(* IEC 61131-3 sources: TetherPLC/tests/ops/cases, 40 files *)

(* ---- o01_debounce.st ---- *)
// o01_debounce.st — FB_AtcDebounce: OnTime=0.3 s sets Q, OffTime=0.2 s
// resets it, ct=0.1 s/scan. D high at n=1 -> Q at n=3 (0.3 s).
// D low at n=6 -> Q clears at n=7 (0.2 s). ET counts since change.
// Sticky bits -> flags %QB0: b0 Q set, b1 Q cleared, b2 ET sane.
PROGRAM O01
VAR
    flags AT %QB0 : BYTE;
    ok0, ok1, ok2 : BOOL;
    deb : FB_AtcDebounce;
    d : BOOL;
    n : DINT;
END_VAR
    n := n + 1;
    IF n = 1 THEN d := TRUE; END_IF;
    IF n = 6 THEN d := FALSE; END_IF;
    deb(D := d, OnTime := 0.3, OffTime := 0.2, CycleTime := 0.1);
    IF n >= 3 AND n < 6 AND deb.Q THEN ok0 := TRUE; END_IF;
    IF n >= 7 AND NOT deb.Q AND n < 30 THEN ok1 := TRUE; END_IF;
    IF n >= 10 AND n < 30 AND deb.ET > 0.05 THEN ok2 := TRUE; END_IF;
    flags := 0;
    IF ok0 THEN flags := flags + 1; END_IF;
    IF ok1 THEN flags := flags + 2; END_IF;
    IF ok2 THEN flags := flags + 4; END_IF;
END_PROGRAM

(* ---- o02_alarm.st ---- *)
// o02_alarm.st — FB_AtcAlarm: Cond edge latches Unacked (survives
// Cond clear), Ack clears it, Shelve suppresses Active for
// ShelveTime s, FirstOut respects HigherPriActive.
//   n=1 Cond up   -> Active+Unacked, FirstOut (no higher pri)
//   n=2 Cond down -> Unacked stays, Active off
//   n=3 Ack       -> Unacked off
//   n=4 Cond up   -> edge again (ack still held -> net unacked off)
//   n=5 Shelve 1s -> Active off, Shelved on
//   n=6..13 shelf window: alm2 (same cond, no shelve, higher-pri =
//        alm.Active=FALSE) -> FirstOut TRUE while alm suppressed
//   n=15+ shelf expires -> alm Active back -> alm2 FirstOut off
// Sticky: b0 unacked latch, b1 ack clears, b2 shelve works,
// b3 shelf expiry restores, b4 firstout suppression.
PROGRAM O02
VAR
    flags AT %QB0 : BYTE;
    ok0, ok1, ok2, ok3, ok4 : BOOL;
    alm : FB_AtcAlarm;
    alm2 : FB_AtcAlarm;
    cond, ack, shelve : BOOL;
    n : DINT;
END_VAR
    n := n + 1;
    IF n = 1 THEN cond := TRUE; END_IF;
    IF n = 2 THEN cond := FALSE; END_IF;
    IF n = 3 THEN ack := TRUE; END_IF;
    IF n = 4 THEN cond := TRUE; END_IF;
    IF n = 5 THEN shelve := TRUE; ack := FALSE; END_IF;
    IF n = 6 THEN shelve := FALSE; END_IF;
    alm(Cond := cond, Ack := ack, Shelve := shelve,
        ShelveTime := 1.0, HigherPriActive := FALSE,
        CycleTime := 0.1);
    alm2(Cond := cond, Ack := FALSE, Shelve := FALSE,
         ShelveTime := 1.0, HigherPriActive := alm.Active,
         CycleTime := 0.1);
    // b0: unacked latched at n=2 even though cond cleared
    IF n = 2 AND alm.Unacked AND NOT alm.Active THEN ok0 := TRUE; END_IF;
    // b1: ack at n=3 cleared unacked
    IF n = 3 AND NOT alm.Unacked THEN ok1 := TRUE; END_IF;
    // b2: shelved at n=6 — cond up but Active suppressed
    IF n = 6 AND alm.Shelved AND NOT alm.Active AND alm.ShelfET > 0.5
       THEN ok2 := TRUE; END_IF;
    // b3: shelf expired -> Active again while cond still up
    IF n >= 15 AND alm.Active AND NOT alm.Shelved THEN ok3 := TRUE; END_IF;
    // b4: during shelf window alm2 is the first-out (alm suppressed)
    IF n = 8 AND alm2.FirstOut AND NOT alm.Active THEN ok4 := TRUE; END_IF;
    flags := 0;
    IF ok0 THEN flags := flags + 1; END_IF;
    IF ok1 THEN flags := flags + 2; END_IF;
    IF ok2 THEN flags := flags + 4; END_IF;
    IF ok3 THEN flags := flags + 8; END_IF;
    IF ok4 THEN flags := flags + 16; END_IF;
END_PROGRAM

(* ---- o03_hourmeter.st ---- *)
// o03_hourmeter.st — FB_AtcHourMeter: ct=3600 s/scan so each scan is
// one hour. Run scans 1-3 -> Hours=3.0, Preset=2.5 -> Alarm + Pct=120.
// Run off at n=4 (hours hold), Reset at n=6 -> zeroed.
// Sticky: b0 hours accumulate, b1 alarm+pct, b2 reset clears.
PROGRAM O03
VAR
    flags AT %QB0 : BYTE;
    ok0, ok1, ok2 : BOOL;
    hm : FB_AtcHourMeter;
    run, rst : BOOL;
    n : DINT;
END_VAR
    n := n + 1;
    run := n <= 3;
    IF n = 6 THEN rst := TRUE; END_IF;
    hm(Run := run, CycleTime := 3600.0, Preset := 2.5, Reset := rst);
    IF n = 3 AND hm.Hours > 2.9 AND hm.Hours < 3.1 THEN ok0 := TRUE; END_IF;
    IF n = 4 AND hm.Alarm AND hm.Pct > 110.0 THEN ok1 := TRUE; END_IF;
    IF n = 7 AND hm.Hours = 0.0 AND NOT hm.Alarm THEN ok2 := TRUE; END_IF;
    flags := 0;
    IF ok0 THEN flags := flags + 1; END_IF;
    IF ok1 THEN flags := flags + 2; END_IF;
    IF ok2 THEN flags := flags + 4; END_IF;
END_PROGRAM

(* ---- o04_oee.st ---- *)
// o04_oee.st — FB_AtcOee: ct=3600 -> 1 h/scan. Planned+Running all
// scans; IdealCycle=10 s. GoodPart pulse n=1, TotalPart pulses n=1,2.
// After n=2: A=100, P=10/(2*3600)*100=0.139, Q=50, OEE~0.069.
// n=8 Reset -> all counters zero, A back to 0 (no plan time).
// Sticky: b0 availability 100, b1 quality 50, b2 perf in band,
// b3 oee in band, b4 reset.
PROGRAM O04
VAR
    flags AT %QB0 : BYTE;
    ok0, ok1, ok2, ok3, ok4 : BOOL;
    oee : FB_AtcOee;
    good, tot, rst : BOOL;
    n : DINT;
END_VAR
    n := n + 1;
    good := n = 1;
    tot := n <= 2;
    rst := n = 8;
    oee(Planned := TRUE, Running := TRUE, IdealCycle := 10.0,
        GoodPart := good, TotalPart := tot, Reset := rst,
        CycleTime := 3600.0);
    IF n = 2 AND oee.Availability > 99.9 THEN ok0 := TRUE; END_IF;
    IF n = 2 AND oee.Quality > 49.9 AND oee.Quality < 50.1
       THEN ok1 := TRUE; END_IF;
    IF n = 2 AND oee.Performance > 0.1 AND oee.Performance < 0.2
       THEN ok2 := TRUE; END_IF;
    IF n = 2 AND oee.OEE > 0.05 AND oee.OEE < 0.09 THEN ok3 := TRUE; END_IF;
    IF n = 9 AND oee.GoodCount = 0 AND oee.TotalCount = 0
       AND oee.PlannedH < 1.5 THEN ok4 := TRUE; END_IF;
    flags := 0;
    IF ok0 THEN flags := flags + 1; END_IF;
    IF ok1 THEN flags := flags + 2; END_IF;
    IF ok2 THEN flags := flags + 4; END_IF;
    IF ok3 THEN flags := flags + 8; END_IF;
    IF ok4 THEN flags := flags + 16; END_IF;
END_PROGRAM

(* ---- o05_sensorcheck.st ---- *)
// o05_sensorcheck.st — FB_AtcSensorCheck: Min=0 Max=100 MaxRate=50
// EU/s StuckBand=0.5 StuckTime=1.0 ct=0.1.
//   n=1  In=50 init (no rate/frozen yet)
//   n=2.. In=50 frozen -> Reason=3 Bad latches ~n=6 (0.5 s)
//   n=12 In=150 -> range Reason=1
//   n=13 In=50 -> in range again; Bad stays latched (Reason=1 latched)
//   n=14 Reset -> Bad/Reason clear
//   n=15 In=80 jump +30 in 0.1 s -> rate 300>50 Reason=2
//   n=16 In=80.4 (within band) frozen resumes
// Sticky: b0 stuck reason3, b1 range reason1, b2 bad latched,
// b3 rate reason2, b4 reset clears.
PROGRAM O05
VAR
    flags AT %QB0 : BYTE;
    ok0, ok1, ok2, ok3, ok4 : BOOL;
    sc : FB_AtcSensorCheck;
    inp : LREAL;
    rst : BOOL;
    n : DINT;
END_VAR
    n := n + 1;
    inp := 50.0;
    IF n = 1 THEN inp := 50.0; END_IF;
    IF n = 12 THEN inp := 150.0; END_IF;
    IF n = 13 THEN inp := 50.0; END_IF;
    rst := n = 14 OR n = 16;
    IF n = 15 THEN inp := 80.0; END_IF;
    IF n >= 16 THEN inp := 80.4; END_IF;
    // n=15 rate violation latches Bad; n=16 resets to check recovery
    sc(In := inp, Min := 0.0, Max := 100.0, MaxRate := 50.0,
       StuckBand := 0.5, StuckTime := 0.5, Reset := rst,
       CycleTime := 0.1);
    IF n >= 7 AND n <= 11 AND sc.Reason = 3 AND sc.Bad THEN ok0 := TRUE; END_IF;
    IF n = 12 AND sc.Reason = 1 THEN ok1 := TRUE; END_IF;
    IF n = 13 AND sc.Bad AND NOT sc.Ok THEN ok2 := TRUE; END_IF;
    IF n = 15 AND sc.Reason = 2 THEN ok3 := TRUE; END_IF;
    IF n = 16 AND NOT sc.Bad AND sc.Ok AND sc.Reason = 0
       THEN ok4 := TRUE; END_IF;
    flags := 0;
    IF ok0 THEN flags := flags + 1; END_IF;
    IF ok1 THEN flags := flags + 2; END_IF;
    IF ok2 THEN flags := flags + 4; END_IF;
    IF ok3 THEN flags := flags + 8; END_IF;
    IF ok4 THEN flags := flags + 16; END_IF;
END_PROGRAM

(* ---- o06_seq.st ---- *)
// o06_seq.st — FB_AtcSeq drum sequencer, ct=0.1.
//   step1 TIME=0.5 NEXT=2 EV=1 ; step2 TIME=0 (wait StepDone)
//   NEXT=3 EV=2 ; step3 TIME=0.5 NEXT=0 EV=4
//   n=1 RUN -> step1; StepTime hits 0.5 at n=6 -> step2
//   n=8 StepDone pulse -> step3; hits 0.5 at n=13 -> NEXT=0
//   n=14 Done, Busy off.
// Sticky: b0 step1 active, b1 step2 reached, b2 step3 via StepDone,
// b3 Done+not Busy, b4 EV of step3 seen.
PROGRAM O06
VAR
    flags AT %QB0 : BYTE;
    ok0, ok1, ok2, ok3, ok4 : BOOL;
    sq : FB_AtcSeq;
    run, sdone : BOOL;
    n : DINT;
END_VAR
    n := n + 1;
    // segment table written member-wise (aggregates can't bind)
    IF n = 1 THEN
        sq.STEPS[1].TIME := 0.5; sq.STEPS[1].NEXT := 2;
        sq.STEPS[1].EV := 1;
        sq.STEPS[2].TIME := 0.0; sq.STEPS[2].NEXT := 3;
        sq.STEPS[2].EV := 2;
        sq.STEPS[3].TIME := 0.5; sq.STEPS[3].NEXT := 0;
        sq.STEPS[3].EV := 4;
    END_IF;
    IF n = 1 THEN run := TRUE; END_IF;
    IF n = 8 THEN sdone := TRUE; END_IF;
    IF n = 9 THEN sdone := FALSE; END_IF;
    sq(NUM_STEPS := 3, RUN := run, HOLD := FALSE,
       RESET := FALSE, StepDone := sdone, CycleTime := 0.1);
    IF n = 3 AND sq.StepIdx = 1 AND sq.Busy THEN ok0 := TRUE; END_IF;
    IF n = 7 AND sq.StepIdx = 2 THEN ok1 := TRUE; END_IF;
    IF n = 9 AND sq.StepIdx = 3 THEN ok2 := TRUE; END_IF;
    IF n >= 14 AND sq.Done AND NOT sq.Busy THEN ok3 := TRUE; END_IF;
    IF n = 10 AND sq.EV = 4 THEN ok4 := TRUE; END_IF;
    flags := 0;
    IF ok0 THEN flags := flags + 1; END_IF;
    IF ok1 THEN flags := flags + 2; END_IF;
    IF ok2 THEN flags := flags + 4; END_IF;
    IF ok3 THEN flags := flags + 8; END_IF;
    IF ok4 THEN flags := flags + 16; END_IF;
END_PROGRAM

(* ---- o07_andon.st ---- *)
// o07_andon.st — FB_AtcAndon: combinational priority mapping.
//   n=1 Run        -> Green
//   n=2 +Warning   -> Amber, Green off
//   n=3 +Alarm     -> Red+Buzz, Amber still (Warn held)
//   n=5 all clear +Changeover -> Blue, Green suppressed
//   n=6 Maintenance -> Amber (no Run)
// Sticky bits per output seen in its expected phase.
PROGRAM O07
VAR
    flags AT %QB0 : BYTE;
    ok0, ok1, ok2, ok3, ok4 : BOOL;
    an : FB_AtcAndon;
    n : DINT;
END_VAR
    n := n + 1;
    an(Run := n <= 4 OR n = 5, Warning := n = 2 OR n = 3,
       Alarm := n = 3, Fault := FALSE,
       Maintenance := n = 6, Changeover := n = 5);
    IF n = 1 AND an.Green AND NOT an.Red AND NOT an.Amber
       THEN ok0 := TRUE; END_IF;
    IF n = 2 AND an.Amber AND NOT an.Green AND NOT an.Red
       THEN ok1 := TRUE; END_IF;
    IF n = 3 AND an.Red AND an.Buzzer AND an.Amber
       THEN ok2 := TRUE; END_IF;
    IF n = 5 AND an.Blue AND NOT an.Green AND NOT an.Red
       THEN ok3 := TRUE; END_IF;
    IF n = 6 AND an.Amber AND NOT an.Green THEN ok4 := TRUE; END_IF;
    flags := 0;
    IF ok0 THEN flags := flags + 1; END_IF;
    IF ok1 THEN flags := flags + 2; END_IF;
    IF ok2 THEN flags := flags + 4; END_IF;
    IF ok3 THEN flags := flags + 8; END_IF;
    IF ok4 THEN flags := flags + 16; END_IF;
END_PROGRAM

(* ---- o08_recipe.st ---- *)
// o08_recipe.st — FB_AtcRecipe: 16x16 LREAL store.
//   n=1 write (set2,param3)=42.5 ; n=2 read -> 42.5 Valid
//   n=3 write (set5,param0)=7.0  ; n=4 read -> 7.0 (same instance,
//        different addressing — proves set/param independence)
//   n=5 Clear -> n=6 read -> 0.0
//   n=7 invalid read (set99) -> Valid FALSE Val 0
// Sticky: b0 roundtrip, b1 set independence, b2 clear, b3 invalid.
PROGRAM O08
VAR
    flags AT %QB0 : BYTE;
    ok0, ok1, ok2, ok3 : BOOL;
    rc : FB_AtcRecipe;
    wrSet, wrPar, rdSet, rdPar : DINT;
    wrVal : LREAL;
    n : DINT;
END_VAR
    n := n + 1;
    // default: read back set2 param3; write set2 param3 = 42.5
    rdSet := 2; rdPar := 3;
    wrSet := 2; wrPar := 3; wrVal := 42.5;
    IF n = 1 OR n = 3 THEN
        // n=3 retargets the write to set5 param0 = 7.0
        IF n = 3 THEN
            wrSet := 5; wrPar := 0; wrVal := 7.0;
        END_IF;
    END_IF;
    IF n = 4 OR n = 6 THEN rdSet := 5; rdPar := 0; END_IF;
    IF n = 7 THEN rdSet := 99; rdPar := 0; END_IF;
    rc(WrSet := wrSet, WrParam := wrPar, WrVal := wrVal,
       WrStrobe := (n = 1) OR (n = 3),
       RdSet := rdSet, RdParam := rdPar, Clear := n = 5);
    IF n = 2 AND rc.Val > 42.4 AND rc.Val < 42.6 AND rc.Valid
       THEN ok0 := TRUE; END_IF;
    IF n = 4 AND rc.Val > 6.9 AND rc.Val < 7.1 AND rc.Valid
       THEN ok1 := TRUE; END_IF;
    IF n = 6 AND rc.Val = 0.0 AND rc.Valid THEN ok2 := TRUE; END_IF;
    IF n = 7 AND NOT rc.Valid AND rc.Val = 0.0 THEN ok3 := TRUE; END_IF;
    flags := 0;
    IF ok0 THEN flags := flags + 1; END_IF;
    IF ok1 THEN flags := flags + 2; END_IF;
    IF ok2 THEN flags := flags + 4; END_IF;
    IF ok3 THEN flags := flags + 8; END_IF;
END_PROGRAM

(* ---- o09_onoff.st ---- *)
// o09_onoff.st — FB_AtcOnOff hysteresis. SP=20 Hyst=4 -> band 18..22.
// pv=10 on-side n<=3, pv=20 inside n=4..6 (holds), pv=23 off-side n>=7.
// Sticky: b0 on, b1 held in deadband, b2 off.
PROGRAM O09
VAR
    flags AT %QB0 : BYTE;
    ok0, ok1, ok2 : BOOL;
    oo : FB_AtcOnOff;
    pv : LREAL;
    n : DINT;
END_VAR
    n := n + 1;
    pv := 23.0;
    IF n <= 3 THEN pv := 10.0; END_IF;
    IF n >= 4 AND n <= 6 THEN pv := 20.0; END_IF;
    oo(PV := pv, SP := 20.0, Hyst := 4.0, Enable := TRUE);
    IF n = 3 AND oo.Out THEN ok0 := TRUE; END_IF;
    IF n = 5 AND oo.Out THEN ok1 := TRUE; END_IF;
    IF n = 8 AND NOT oo.Out THEN ok2 := TRUE; END_IF;
    flags := 0;
    IF ok0 THEN flags := flags + 1; END_IF;
    IF ok1 THEN flags := flags + 2; END_IF;
    IF ok2 THEN flags := flags + 4; END_IF;
END_PROGRAM

(* ---- o10_permissive.st ---- *)
// o10_permissive.st — FB_AtcPermissive 8-input AND chain.
// all true n<=2; P3+P5 low n=3..4; only P8 low n=5..6; all n>=7.
// Sticky: b0 permit clear, b1 first-deny=3 mask=20, b2 first-deny=8
// mask=128.
PROGRAM O10
VAR
    flags AT %QB0 : BYTE;
    ok0, ok1, ok2 : BOOL;
    pm : FB_AtcPermissive;
    p3, p5, p8 : BOOL;
    n : DINT;
END_VAR
    n := n + 1;
    p3 := TRUE; p5 := TRUE; p8 := TRUE;
    IF n >= 3 AND n <= 4 THEN p3 := FALSE; p5 := FALSE; END_IF;
    IF n >= 5 AND n <= 6 THEN p8 := FALSE; END_IF;
    pm(P1 := TRUE, P2 := TRUE, P3 := p3, P4 := TRUE,
       P5 := p5, P6 := TRUE, P7 := TRUE, P8 := p8);
    IF n = 2 AND pm.Permit AND pm.DenyMask = 0 THEN ok0 := TRUE; END_IF;
    IF n = 4 AND NOT pm.Permit AND pm.FirstDeny = 3
       AND pm.DenyMask = 20 THEN ok1 := TRUE; END_IF;
    IF n = 6 AND pm.FirstDeny = 8 AND pm.DenyMask = 128
       THEN ok2 := TRUE; END_IF;
    flags := 0;
    IF ok0 THEN flags := flags + 1; END_IF;
    IF ok1 THEN flags := flags + 2; END_IF;
    IF ok2 THEN flags := flags + 4; END_IF;
END_PROGRAM

(* ---- o11_mode.st ---- *)
// o11_mode.st — FB_AtcMode arbitration, priority jog>maint>man>auto.
// n=1..2 auto; n=3..4 man+auto; n=5..6 jog+man+maint; n=7..8 maint;
// n>=9 none. Sticky: b0 auto, b1 man beats auto, b2 jog top,
// b3 maint alone, b4 off-transition Changed.
PROGRAM O11
VAR
    flags AT %QB0 : BYTE;
    ok0, ok1, ok2, ok3, ok4 : BOOL;
    md : FB_AtcMode;
    ra, rm, rj, rh : BOOL;
    n : DINT;
END_VAR
    n := n + 1;
    ra := n <= 4;
    rm := n >= 3 AND n <= 6;
    rj := n >= 5 AND n <= 6;
    rh := n >= 5 AND n <= 8;
    md(ReqAuto := ra, ReqMan := rm, ReqJog := rj, ReqMaint := rh);
    IF n = 2 AND md.Mode = 1 AND md.Auto THEN ok0 := TRUE; END_IF;
    IF n = 4 AND md.Mode = 2 AND md.Man AND NOT md.Auto
       THEN ok1 := TRUE; END_IF;
    IF n = 6 AND md.Mode = 3 AND md.Jog THEN ok2 := TRUE; END_IF;
    IF n = 8 AND md.Mode = 4 AND md.Maint THEN ok3 := TRUE; END_IF;
    IF n = 9 AND md.Mode = 0 AND md.Changed THEN ok4 := TRUE; END_IF;
    flags := 0;
    IF ok0 THEN flags := flags + 1; END_IF;
    IF ok1 THEN flags := flags + 2; END_IF;
    IF ok2 THEN flags := flags + 4; END_IF;
    IF ok3 THEN flags := flags + 8; END_IF;
    IF ok4 THEN flags := flags + 16; END_IF;
END_PROGRAM

(* ---- o12_jog.st ---- *)
// o12_jog.st — FB_AtcJog deadman + anti-run timeout, ct=0.1 MaxOn=0.3.
// En+Dir=+1 n=2..5: ET hits 0.3 at n=4 -> Out drops, TimedOut latches
// while En held; n=6 En released -> clears.
// Sticky: b0 jogging, b1 timed out, b2 released-clear.
PROGRAM O12
VAR
    flags AT %QB0 : BYTE;
    ok0, ok1, ok2 : BOOL;
    jg : FB_AtcJog;
    en : BOOL;
    n : DINT;
END_VAR
    n := n + 1;
    en := n >= 2 AND n <= 5;
    jg(DirIn := 1, En := en, MaxOn := 0.3, CycleTime := 0.1);
    IF n = 3 AND jg.Out AND jg.Dir = 1 AND NOT jg.TimedOut
       THEN ok0 := TRUE; END_IF;
    IF n = 5 AND NOT jg.Out AND jg.TimedOut THEN ok1 := TRUE; END_IF;
    IF n = 7 AND NOT jg.TimedOut AND NOT jg.Out THEN ok2 := TRUE; END_IF;
    flags := 0;
    IF ok0 THEN flags := flags + 1; END_IF;
    IF ok1 THEN flags := flags + 2; END_IF;
    IF ok2 THEN flags := flags + 4; END_IF;
END_PROGRAM

(* ---- o13_watchdog.st ---- *)
// o13_watchdog.st — FB_AtcWatchdog heartbeat, ct=0.1 Timeout=0.25.
// Kick pulses n=1,3,5,7 then stops: ET grows past 0.25 at n=10.
// Sticky: b0 ok between kicks, b1 ok near timeout, b2 err latched.
PROGRAM O13
VAR
    flags AT %QB0 : BYTE;
    ok0, ok1, ok2 : BOOL;
    wd : FB_AtcWatchdog;
    kick : BOOL;
    n : DINT;
END_VAR
    n := n + 1;
    kick := n = 1 OR n = 3 OR n = 5 OR n = 7;
    wd(Kick := kick, Timeout := 0.25, CycleTime := 0.1,
       Reset := FALSE);
    IF n = 6 AND wd.OK AND wd.ET > 0.05 AND wd.ET < 0.15
       THEN ok0 := TRUE; END_IF;
    IF n = 9 AND wd.OK AND wd.ET > 0.15 THEN ok1 := TRUE; END_IF;
    IF n = 11 AND wd.Err AND NOT wd.OK THEN ok2 := TRUE; END_IF;
    flags := 0;
    IF ok0 THEN flags := flags + 1; END_IF;
    IF ok1 THEN flags := flags + 2; END_IF;
    IF ok2 THEN flags := flags + 4; END_IF;
END_PROGRAM

(* ---- o14_blinker.st ---- *)
// o14_blinker.st — FB_AtcBlinker Rate=2Hz Duty=0.5 ct=0.1 -> 5-scan
// period, Q on ~first half. frac sequence 0.2,0.4,0.6,0.8,wrap.
// Sample away from the 0.5 boundary for float safety.
// Sticky: b0 on, b1 off, b2 wrapped-on, b3 off again.
PROGRAM O14
VAR
    flags AT %QB0 : BYTE;
    ok0, ok1, ok2, ok3 : BOOL;
    bl : FB_AtcBlinker;
    n : DINT;
END_VAR
    n := n + 1;
    bl(En := TRUE, Rate := 2.0, Duty := 0.5, CycleTime := 0.1);
    IF n = 1 AND bl.Q THEN ok0 := TRUE; END_IF;
    IF n = 3 AND NOT bl.Q THEN ok1 := TRUE; END_IF;
    IF n = 6 AND bl.Q THEN ok2 := TRUE; END_IF;
    IF n = 8 AND NOT bl.Q THEN ok3 := TRUE; END_IF;
    flags := 0;
    IF ok0 THEN flags := flags + 1; END_IF;
    IF ok1 THEN flags := flags + 2; END_IF;
    IF ok2 THEN flags := flags + 4; END_IF;
    IF ok3 THEN flags := flags + 8; END_IF;
END_PROGRAM

(* ---- o15_totalizer.st ---- *)
// o15_totalizer.st — FB_AtcTotalizer Rate=2 K=3 ct=0.1 -> +0.6/scan.
// Reset at n=4 zeroes; accumulation resumes.
// Sticky: b0 accumulates, b1 reset, b2 resumes.
PROGRAM O15
VAR
    flags AT %QB0 : BYTE;
    ok0, ok1, ok2 : BOOL;
    tz : FB_AtcTotalizer;
    rst : BOOL;
    n : DINT;
END_VAR
    n := n + 1;
    rst := n = 4;
    tz(Rate := 2.0, K := 3.0, CycleTime := 0.1, Reset := rst);
    IF n = 3 AND tz.Total > 1.7 AND tz.Total < 1.9
       THEN ok0 := TRUE; END_IF;
    IF n = 4 AND tz.Total = 0.0 THEN ok1 := TRUE; END_IF;
    IF n = 6 AND tz.Total > 1.1 AND tz.Total < 1.3
       THEN ok2 := TRUE; END_IF;
    flags := 0;
    IF ok0 THEN flags := flags + 1; END_IF;
    IF ok1 THEN flags := flags + 2; END_IF;
    IF ok2 THEN flags := flags + 4; END_IF;
END_PROGRAM

(* ---- o16_avg.st ---- *)
// o16_avg.st — FB_AtcAvg N=3 window over av=n*10.
// n=3 avg 20; n=4 window {40,20,30} avg 30; n=5 {40,50,30} avg 40.
// Sticky: b0/b1/b2 window means.
PROGRAM O16
VAR
    flags AT %QB0 : BYTE;
    ok0, ok1, ok2 : BOOL;
    av2 : FB_AtcAvg;
    av : LREAL;
    n : DINT;
END_VAR
    n := n + 1;
    av := n * 10.0;
    av2(In := av, N := 3);
    IF n = 3 AND av2.Avg > 19.9 AND av2.Avg < 20.1
       AND av2.Count = 3 THEN ok0 := TRUE; END_IF;
    IF n = 4 AND av2.Avg > 29.9 AND av2.Avg < 30.1
       THEN ok1 := TRUE; END_IF;
    IF n = 5 AND av2.Avg > 39.9 AND av2.Avg < 40.1
       THEN ok2 := TRUE; END_IF;
    flags := 0;
    IF ok0 THEN flags := flags + 1; END_IF;
    IF ok1 THEN flags := flags + 2; END_IF;
    IF ok2 THEN flags := flags + 4; END_IF;
END_PROGRAM

(* ---- o17_demand.st ---- *)
// o17_demand.st — FB_AtcDemand Window=0.25 ct=0.1 -> n=2 samples.
// pw=n*10. n=3 window {30,20} -> 25; n=5 {50,40} -> 45;
// n=6 Reset; n=7 single sample 70 -> 70.
// Sticky: b0/b1 windowed mean, b2 post-reset restart.
PROGRAM O17
VAR
    flags AT %QB0 : BYTE;
    ok0, ok1, ok2 : BOOL;
    dm : FB_AtcDemand;
    rst : BOOL;
    pw : LREAL;
    n : DINT;
END_VAR
    n := n + 1;
    pw := n * 10.0;
    rst := n = 6;
    dm(Power := pw, Window := 0.25, CycleTime := 0.1,
       Reset := rst);
    IF n = 3 AND dm.Demand > 24.9 AND dm.Demand < 25.1
       THEN ok0 := TRUE; END_IF;
    IF n = 5 AND dm.Demand > 44.9 AND dm.Demand < 45.1
       THEN ok1 := TRUE; END_IF;
    IF n = 7 AND dm.Demand > 69.9 AND dm.Demand < 70.1
       AND dm.Samples = 1 THEN ok2 := TRUE; END_IF;
    flags := 0;
    IF ok0 THEN flags := flags + 1; END_IF;
    IF ok1 THEN flags := flags + 2; END_IF;
    IF ok2 THEN flags := flags + 4; END_IF;
END_PROGRAM

(* ---- o18_override.st ---- *)
// o18_override.st — FB_AtcOverride manual/auto + release track.
// AutoIn=50 ManIn=80 TrackIn=60; ManEn n=2..4.
// n=5 release scan -> Out=TrackIn=60 Tracking; n>=6 -> AutoIn=50.
// Sticky: b0 manual, b1 release-sync, b2 auto passthrough.
PROGRAM O18
VAR
    flags AT %QB0 : BYTE;
    ok0, ok1, ok2 : BOOL;
    ov : FB_AtcOverride;
    men : BOOL;
    n : DINT;
END_VAR
    n := n + 1;
    men := n >= 2 AND n <= 4;
    ov(AutoIn := 50.0, ManIn := 80.0, ManEn := men,
       TrackIn := 60.0);
    IF n = 3 AND ov.Out = 80.0 THEN ok0 := TRUE; END_IF;
    IF n = 5 AND ov.Tracking AND ov.Out = 60.0 THEN ok1 := TRUE; END_IF;
    IF n = 7 AND NOT ov.Tracking AND ov.Out = 50.0
       THEN ok2 := TRUE; END_IF;
    flags := 0;
    IF ok0 THEN flags := flags + 1; END_IF;
    IF ok1 THEN flags := flags + 2; END_IF;
    IF ok2 THEN flags := flags + 4; END_IF;
END_PROGRAM

(* ---- o19_twohand.st ---- *)
// o19_twohand.st — FB_AtcTwoHand anti-tie-down, ct=0.1 MaxGap=0.5.
// Btn1 n=2..5, Btn2 n=4..7: valid press -> Out while both held.
// Btn1 released n=6 -> Out drops. n=8+ both released -> disarm.
// n=9 Btn1 held alone -> gap expires n=14; Btn2 tap n=15 rejected.
// Sticky: b0 permit, b1 release-drop, b2 disarmed, b3 late-tap reject.
PROGRAM O19
VAR
    flags AT %QB0 : BYTE;
    ok0, ok1, ok2, ok3 : BOOL;
    th : FB_AtcTwoHand;
    b1, b2 : BOOL;
    n : DINT;
END_VAR
    n := n + 1;
    b1 := (n >= 2 AND n <= 5) OR (n >= 9 AND n <= 16);
    b2 := (n >= 4 AND n <= 7) OR n = 15;
    th(Btn1 := b1, Btn2 := b2, MaxGap := 0.5,
       CycleTime := 0.1, Reset := FALSE);
    IF n = 5 AND th.Out AND th.Armed THEN ok0 := TRUE; END_IF;
    IF n = 6 AND NOT th.Out THEN ok1 := TRUE; END_IF;
    IF n = 14 AND NOT th.Armed THEN ok2 := TRUE; END_IF;
    IF n = 16 AND NOT th.Out AND NOT th.Armed THEN ok3 := TRUE; END_IF;
    flags := 0;
    IF ok0 THEN flags := flags + 1; END_IF;
    IF ok1 THEN flags := flags + 2; END_IF;
    IF ok2 THEN flags := flags + 4; END_IF;
    IF ok3 THEN flags := flags + 8; END_IF;
END_PROGRAM

(* ---- o20_shift.st ---- *)
// o20_shift.st — FB_AtcShift: S1 08-12, S2 16-20, S3 overnight 22-04.
// TOD := n*1800 (30 min/scan). Checks shift index, start/end pulses,
// elapsed/remaining, and midnight-wrap continuity of the night shift.
// Sticky bits -> flags %QB0: b0 in-shift idx, b1 ShiftEnd seen,
// b2 ShiftStart seen, b3 elapsed/remaining sane.
PROGRAM O20
VAR
    flags AT %QB0 : BYTE;
    ok0, ok1, ok2, ok3 : BOOL;
    sh : FB_AtcShift;
    tod : LREAL;
    n : DINT;
    endSeen, startSeen : BOOL;
    elOk, remOk : BOOL;
END_VAR
    n := n + 1;
    tod := DINT_TO_LREAL(n) * 1800.0;
    sh(TOD := tod, Enable := TRUE,
       S1Start := 28800.0, S1End := 43200.0,
       S2Start := 57600.0, S2End := 72000.0,
       S3Start := 79200.0, S3End := 14400.0);
    endSeen := endSeen OR sh.ShiftEnd;
    startSeen := startSeen OR sh.ShiftStart;
    // b0: correct shift index across the day (S3 early, S1 mid, S2 eve)
    IF (n <= 7 AND sh.Shift = 3 AND sh.InShift)
       OR (n >= 16 AND n <= 23 AND sh.Shift = 1 AND sh.InShift)
       OR (n >= 32 AND n <= 39 AND sh.Shift = 2 AND sh.InShift)
       OR (n >= 44 AND n <= 55 AND sh.Shift = 3 AND sh.InShift) THEN
        ok0 := TRUE;
    END_IF;
    // b1: left-shift pulse fired at the 04:00, 12:00, 20:00 boundaries
    IF n >= 9 AND endSeen THEN ok1 := TRUE; END_IF;
    // b2: entered-shift pulse fired at 08:00, 16:00, 22:00, and 00:00-wrap
    IF n >= 17 AND startSeen THEN ok2 := TRUE; END_IF;
    // b3: elapsed/remaining sane — n=17 is 30 min into S1;
    // n=50 is 01:00 inside overnight S3 (elapsed 3h, remaining 3h)
    elOk := FALSE; remOk := FALSE;
    IF n = 17 THEN
        IF sh.Elapsed > 1700.0 AND sh.Elapsed < 1900.0
           AND sh.Remaining > 12000.0 AND sh.Remaining < 13200.0 THEN
            elOk := TRUE; remOk := TRUE;
        END_IF;
    END_IF;
    IF n = 50 THEN
        IF sh.Elapsed > 10000.0 AND sh.Elapsed < 11600.0
           AND sh.Remaining > 10000.0 AND sh.Remaining < 11600.0 THEN
            elOk := TRUE; remOk := TRUE;
        END_IF;
    END_IF;
    IF elOk AND remOk THEN ok3 := TRUE; END_IF;
    flags := 0;
    IF ok0 THEN flags := flags + 1; END_IF;
    IF ok1 THEN flags := flags + 2; END_IF;
    IF ok2 THEN flags := flags + 4; END_IF;
    IF ok3 THEN flags := flags + 8; END_IF;
END_PROGRAM

(* ---- o21_defrost.st ---- *)
// o21_defrost.st — FB_AtcDefrost: DefrostEvery=2 s, DefrostTime=0.5 s,
// MinOff=0.5 s, ct=0.1. Cool n=1..19, defrost ~n=20..23, off-delay
// ~n=24..30 (float offT needs an extra scan), cool resumes n=31.
// Door ajar n=30..37: qualified door-time starts n=32 (fridgeOn only
// true from n=31), doorT reaches 0.5 at n=36 -> DoorAlarm latches.
// Ack n=39 clears it. Warm n=42..44 latches TempAlarm at n=44.
// Sticky bits -> flags %QB0: expect 0x1f.
PROGRAM O21
VAR
    flags AT %QB0 : BYTE;
    ok0, ok1, ok2, ok3, ok3b, ok4 : BOOL;
    df : FB_AtcDefrost;
    door, warm, ack : BOOL;
    n : DINT;
END_VAR
    n := n + 1;
    IF n >= 30 AND n <= 37 THEN door := TRUE; ELSE door := FALSE; END_IF;
    IF n >= 42 AND n <= 45 THEN warm := TRUE; ELSE warm := FALSE; END_IF;
    ack := (n = 39);
    df(Enable := TRUE, DoorOpen := door, Warm := warm, Ack := ack,
       DefrostEvery := 2.0, DefrostTime := 0.5, MinOff := 0.5,
       DoorAlarmTime := 0.5, WarmTime := 0.3, CycleTime := 0.1);
    IF (n >= 1 AND n <= 19) OR (n >= 31 AND n <= 33) THEN
        IF df.Fridge THEN ok0 := TRUE; END_IF;
    END_IF;
    IF (n = 21 OR n = 22) AND df.DefrostHeat AND df.InDefrost THEN
        ok1 := TRUE;
    END_IF;
    IF n >= 24 AND df.DefrostCount >= 1 THEN ok2 := TRUE; END_IF;
    IF n >= 36 AND n <= 38 AND df.DoorAlarm THEN ok3 := TRUE; END_IF;
    IF n >= 40 AND n <= 44 AND NOT df.DoorAlarm THEN ok3b := TRUE; END_IF;
    IF n >= 45 AND df.TempAlarm THEN ok4 := TRUE; END_IF;
    flags := 0;
    IF ok0 THEN flags := flags + 1; END_IF;
    IF ok1 THEN flags := flags + 2; END_IF;
    IF ok2 THEN flags := flags + 4; END_IF;
    IF ok3 AND ok3b THEN flags := flags + 8; END_IF;
    IF ok4 THEN flags := flags + 16; END_IF;
END_PROGRAM

(* ---- o22_zonebalance.st ---- *)
// o22_zonebalance.st — FB_AtcZoneBalance: Gain=2, TrimMax=5, RateMax=10
// (1 degC/scan at ct=0.1). MasterErr=3 at n=1 -> want=6 clamps to 5,
// rate-limited ramp reaches 5 by n=5, Sat set. MasterErr=0 at n=10 ->
// ramps down 1/scan, hits 0 at n=14. Disable n=20 -> bumpless reset;
// re-enable n=25 starts at 0 again. Per-scan |dTrim| <= 1.01 always.
// Sticky bits -> flags %QB0: expect 0x1f.
PROGRAM O22
VAR
    flags AT %QB0 : BYTE;
    ok0, ok1, ok2, ok3, ok4 : BOOL;
    zb : FB_AtcZoneBalance;
    err : LREAL;
    en : BOOL;
    n : DINT;
    prev : LREAL;
    dmax : LREAL;
    first : BOOL;
END_VAR
    n := n + 1;
    first := (n = 1);
    IF n = 1 THEN err := 3.0; END_IF;
    IF n = 10 THEN err := 0.0; END_IF;
    en := NOT (n >= 20 AND n <= 24);
    zb(MasterErr := err, Enable := en, Gain := 2.0,
       TrimMax := 5.0, RateMax := 10.0, CycleTime := 0.1);
    // per-scan rate-limit invariant
    IF NOT first THEN
        IF zb.TrimOut - prev > dmax THEN
            dmax := zb.TrimOut - prev;
        END_IF;
        IF prev - zb.TrimOut > dmax THEN
            dmax := prev - zb.TrimOut;
        END_IF;
    END_IF;
    prev := zb.TrimOut;
    IF n >= 6 AND n <= 9 AND zb.TrimOut > 4.9 AND zb.Sat THEN
        ok0 := TRUE;
    END_IF;
    IF n >= 6 AND n <= 9 AND zb.Sat THEN ok1 := TRUE; END_IF;
    IF n = 11 AND zb.TrimOut > 2.9 AND zb.TrimOut < 3.1 THEN
        ok2 := TRUE;
    END_IF;
    IF n >= 21 AND n <= 24 AND zb.TrimOut = 0.0 THEN ok3 := TRUE; END_IF;
    IF n = 30 AND zb.TrimOut < 0.2 THEN ok4 := TRUE; END_IF;
    flags := 0;
    IF ok0 THEN flags := flags + 1; END_IF;
    IF ok1 THEN flags := flags + 2; END_IF;
    IF ok2 THEN flags := flags + 4; END_IF;
    IF ok3 THEN flags := flags + 8; END_IF;
    IF ok4 AND dmax <= 1.01 THEN flags := flags + 16; END_IF;
END_PROGRAM

(* ---- o23_endpoint.st ---- *)
// o23_endpoint.st — FB_AtcEndpoint: Execute at n=1, SettleTime=0.5,
// SampleTime=1.0, MaxRise=10/s, ct=0.1. Pressure ramps 50/s during
// the sample window -> RiseRate ~500 -> Result=2 (wet). Checks valve
// isolation, testing flag, wet classification, valve reopen, rate.
// Sticky bits -> flags %QB0: expect 0x1f.
PROGRAM O23
VAR
    flags AT %QB0 : BYTE;
    ok0, ok1, ok2, ok3, ok4 : BOOL;
    ep : FB_AtcEndpoint;
    p : LREAL;
    n : DINT;
    ex : BOOL;
END_VAR
    n := n + 1;
    ex := (n = 1);
    // flat 100 during settle; +50/s ramp once sampling starts (n>5)
    IF n <= 5 THEN p := 100.0;
    ELSE p := 100.0 + DINT_TO_LREAL(n - 5) * 50.0; END_IF;
    ep(Execute := ex, Pressure := p,
       SettleTime := 0.5, SampleTime := 1.0, MaxRise := 10.0,
       CycleTime := 0.1, Reset := FALSE);
    // valve isolated during settle+sample (st 1,2 -> n=2..15)
    IF n >= 3 AND n <= 14 AND NOT ep.ValveCmd THEN ok0 := TRUE; END_IF;
    IF n = 10 AND ep.Testing THEN ok1 := TRUE; END_IF;
    IF n >= 16 AND ep.Result = 2 THEN ok2 := TRUE; END_IF;
    IF n >= 16 AND ep.ValveCmd AND NOT ep.Testing THEN ok3 := TRUE; END_IF;
    IF n >= 16 AND ep.RiseRate > 100.0 THEN ok4 := TRUE; END_IF;
    flags := 0;
    IF ok0 THEN flags := flags + 1; END_IF;
    IF ok1 THEN flags := flags + 2; END_IF;
    IF ok2 THEN flags := flags + 4; END_IF;
    IF ok3 THEN flags := flags + 8; END_IF;
    IF ok4 THEN flags := flags + 16; END_IF;
END_PROGRAM

(* ---- o24_leadlag.st ---- *)
// o24_leadlag.st — FB_AtcLeadLag: 3 units, StageDelay=0.5 s, ct=0.1.
// Stage changes step ONE unit per StageDelay. dem=2 n=11..30:
// onT 0->1 n=11 sel={1}; 1->2 n=16 re-picks least hours -> {2,3}
// (stage1 accrued 0.5 s, 2&3 zero). dem=0 n=31..50: onT 2->1 n=31
// sel={1} (least hrs), 1->0 n=36. dem=1 n=51..60: onT=1 sel={1}
// (1.0 s vs 1.5 s on 2&3). flags %QB0: expect 0x3f.
PROGRAM O24
VAR
    flags AT %QB0 : BYTE;
    ok0, ok1, ok2, ok3, ok4, ok5 : BOOL;
    ll : FB_AtcLeadLag;
    n : DINT;
    dem : LREAL;
END_VAR
    n := n + 1;
    dem := 0.0;
    IF n >= 11 AND n <= 30 THEN dem := 2.0; END_IF;
    IF n >= 51 THEN dem := 1.0; END_IF;
    ll(Demand := dem, NumUnits := 3, StageDelay := 0.5,
       Enable := TRUE, CycleTime := 0.1, Reset := FALSE);
    IF n >= 5 AND n <= 10 AND ll.NumOn = 0 THEN ok0 := TRUE; END_IF;
    IF n >= 12 AND n <= 14 AND ll.NumOn = 1 AND ll.Stage[1]
        AND NOT ll.Stage[2] AND NOT ll.Stage[3] THEN
        ok1 := TRUE;
    END_IF;
    IF n >= 25 AND n <= 30 AND ll.NumOn = 2 AND ll.Stage[2]
        AND ll.Stage[3] AND NOT ll.Stage[1] AND ll.LeadIdx = 2 THEN
        ok2 := TRUE;
    END_IF;
    IF n >= 33 AND n <= 35 AND ll.NumOn = 1 THEN ok3 := TRUE; END_IF;
    IF n >= 40 AND n <= 50 AND ll.NumOn = 0 THEN ok4 := TRUE; END_IF;
    IF n >= 55 AND n <= 60 AND ll.NumOn = 1 AND ll.Stage[1]
        AND ll.LeadIdx = 1 AND NOT ll.Stage[2] AND NOT ll.Stage[3]
    THEN
        ok5 := TRUE;
    END_IF;
    flags := 0;
    IF ok0 THEN flags := flags + 1; END_IF;
    IF ok1 THEN flags := flags + 2; END_IF;
    IF ok2 THEN flags := flags + 4; END_IF;
    IF ok3 THEN flags := flags + 8; END_IF;
    IF ok4 THEN flags := flags + 16; END_IF;
    IF ok5 THEN flags := flags + 32; END_IF;
END_PROGRAM

(* ---- o25_toollife.st ---- *)
// o25_toollife.st — FB_AtcToolLife: LifeLimit=20, WarnPct=80,
// Cycle pulses every even n, Enable while n<45. Cycles hit 16 (80%)
// at n=32 -> Warn; 20 at n=40 -> Due. Reset n=45 clears.
// flags %QB0: expect 0x3f.
PROGRAM O25
VAR
    flags AT %QB0 : BYTE;
    ok0, ok1, ok2, ok3, ok4, ok5 : BOOL;
    tl : FB_AtcToolLife;
    n : DINT;
    cyc : BOOL;
END_VAR
    n := n + 1;
    cyc := (n MOD 2) = 0;
    tl(Cycle := cyc, Enable := (n < 45), LifeLimit := 20,
       WarnPct := 80.0, CycleTime := 0.1, Reset := (n = 45));
    IF n >= 10 AND tl.Cycles >= 5 THEN ok0 := TRUE; END_IF;
    IF n >= 20 AND tl.PctUsed >= 40.0 AND tl.PctUsed < 80.0 THEN
        ok1 := TRUE;
    END_IF;
    IF n >= 33 AND n <= 39 AND tl.Warn AND NOT tl.Due THEN
        ok2 := TRUE;
    END_IF;
    IF n >= 41 AND n <= 44 AND tl.Due THEN ok3 := TRUE; END_IF;
    IF n >= 46 AND tl.Cycles = 0 AND tl.Hours < 0.02 THEN ok4 := TRUE;
    END_IF;
    IF n >= 20 AND n <= 30 AND tl.Hours > 0.0 THEN ok5 := TRUE; END_IF;
    flags := 0;
    IF ok0 THEN flags := flags + 1; END_IF;
    IF ok1 THEN flags := flags + 2; END_IF;
    IF ok2 THEN flags := flags + 4; END_IF;
    IF ok3 THEN flags := flags + 8; END_IF;
    IF ok4 THEN flags := flags + 16; END_IF;
    IF ok5 THEN flags := flags + 32; END_IF;
END_PROGRAM

(* ---- o26_softlimit.st ---- *)
// o26_softlimit.st — FB_AtcSoftLimit: [0,100], Homed from n=11,
// Enable always, Reset n=31. Pos=50 (in), 120 (over n=21..25),
// -10 (under n=26..30), 50 again. PosValid needs Homed; Fault
// latches on first violation, Reset clears.
// flags %QB0: expect 0x3f.
PROGRAM O26
VAR
    flags AT %QB0 : BYTE;
    ok0, ok1, ok2, ok3, ok4, ok5 : BOOL;
    sl : FB_AtcSoftLimit;
    n : DINT;
    pos : LREAL;
    homed : BOOL;
END_VAR
    n := n + 1;
    pos := 50.0;
    IF n >= 21 AND n <= 25 THEN pos := 120.0; END_IF;
    IF n >= 26 AND n <= 30 THEN pos := -10.0; END_IF;
    homed := (n >= 11);
    sl(Pos := pos, MinPos := 0.0, MaxPos := 100.0, Homed := homed,
       Enable := TRUE, Reset := (n = 31));
    IF n >= 5 AND n <= 10 AND NOT sl.PosValid AND sl.NeedHome THEN
        ok0 := TRUE;
    END_IF;
    IF n >= 15 AND n <= 20 AND sl.InWindow AND NOT sl.Fault THEN
        ok1 := TRUE;
    END_IF;
    IF n >= 22 AND n <= 25 AND sl.OverPos AND sl.Fault THEN
        ok2 := TRUE;
    END_IF;
    IF n >= 27 AND n <= 30 AND sl.UnderPos AND sl.Fault THEN
        ok3 := TRUE;
    END_IF;
    IF n >= 32 AND n <= 35 AND NOT sl.Fault AND sl.InWindow THEN
        ok4 := TRUE;
    END_IF;
    IF n >= 12 AND n <= 20 AND sl.PosValid AND NOT sl.NeedHome THEN
        ok5 := TRUE;
    END_IF;
    flags := 0;
    IF ok0 THEN flags := flags + 1; END_IF;
    IF ok1 THEN flags := flags + 2; END_IF;
    IF ok2 THEN flags := flags + 4; END_IF;
    IF ok3 THEN flags := flags + 8; END_IF;
    IF ok4 THEN flags := flags + 16; END_IF;
    IF ok5 THEN flags := flags + 32; END_IF;
END_PROGRAM

(* ---- o27_deviation.st ---- *)
// o27_deviation.st — FB_AtcDeviation: SP=50, Band=5, OnDelay=0.5,
// OffDelay=0.3, ct=0.1. PV=58 n=11..20 (dev 8): Alarm at ~n=15.
// PV=52 n=21..30 (in band): clears ~n=23. PV=54.5 n=31..35 in band.
// PV=60 n=36..45 (dev 10): Alarm again ~n=40.
// flags %QB0: expect 0x3f.
PROGRAM O27
VAR
    flags AT %QB0 : BYTE;
    ok0, ok1, ok2, ok3, ok4, ok5 : BOOL;
    dv : FB_AtcDeviation;
    n : DINT;
    pv : LREAL;
END_VAR
    n := n + 1;
    pv := 50.0;
    IF n >= 11 AND n <= 20 THEN pv := 58.0; END_IF;
    IF n >= 21 AND n <= 30 THEN pv := 52.0; END_IF;
    IF n >= 31 AND n <= 35 THEN pv := 54.5; END_IF;
    IF n >= 36 THEN pv := 60.0; END_IF;
    dv(PV := pv, SP := 50.0, Band := 5.0, OnDelay := 0.5,
       OffDelay := 0.3, Enable := TRUE, CycleTime := 0.1,
       Reset := FALSE);
    IF n >= 12 AND n <= 14 AND dv.Dev AND NOT dv.Alarm THEN
        ok0 := TRUE;
    END_IF;
    IF n >= 17 AND n <= 20 AND dv.Alarm THEN ok1 := TRUE; END_IF;
    IF n = 22 AND dv.Alarm THEN ok2 := TRUE; END_IF;
    IF n >= 25 AND n <= 29 AND NOT dv.Alarm THEN ok3 := TRUE; END_IF;
    IF n >= 41 AND n <= 44 AND dv.Alarm THEN ok4 := TRUE; END_IF;
    IF n >= 17 AND n <= 19 AND dv.ET > 0.2 THEN ok5 := TRUE; END_IF;
    flags := 0;
    IF ok0 THEN flags := flags + 1; END_IF;
    IF ok1 THEN flags := flags + 2; END_IF;
    IF ok2 THEN flags := flags + 4; END_IF;
    IF ok3 THEN flags := flags + 8; END_IF;
    IF ok4 THEN flags := flags + 16; END_IF;
    IF ok5 THEN flags := flags + 32; END_IF;
END_PROGRAM

(* ---- o28_dualchannel.st ---- *)
// o28_dualchannel.st — FB_AtcDualChannel: MismatchTime=0.5, ct=0.1.
// Channels disagree n=11..20: 0.4 s bounce filtered (no fault at
// n=13), 0.5 s at n=15 -> Fault latches; agrees again n=21 but Fault
// stays until Reset n=31. flags %QB0: expect 0x3f.
PROGRAM O28
VAR
    flags AT %QB0 : BYTE;
    ok0, ok1, ok2, ok3, ok4, ok5 : BOOL;
    dc : FB_AtcDualChannel;
    n : DINT;
    i1, i2 : BOOL;
END_VAR
    n := n + 1;
    i1 := TRUE;
    i2 := NOT (n >= 11 AND n <= 20);
    dc(In1 := i1, In2 := i2, MismatchTime := 0.5,
       Enable := TRUE, CycleTime := 0.1, Reset := (n = 31));
    IF n >= 5 AND n <= 10 AND dc.Agree AND dc.Safe THEN ok0 := TRUE;
    END_IF;
    IF n >= 12 AND n <= 14 AND NOT dc.Agree AND NOT dc.Fault THEN
        ok1 := TRUE;
    END_IF;
    IF n >= 16 AND n <= 20 AND dc.Fault AND NOT dc.Safe THEN
        ok2 := TRUE;
    END_IF;
    IF n >= 22 AND n <= 30 AND dc.Agree AND dc.Fault AND NOT dc.Safe
    THEN
        ok3 := TRUE;
    END_IF;
    IF n >= 32 AND n <= 38 AND dc.Safe AND NOT dc.Fault THEN
        ok4 := TRUE;
    END_IF;
    IF n >= 13 AND n <= 14 AND dc.ET > 0.3 THEN ok5 := TRUE; END_IF;
    flags := 0;
    IF ok0 THEN flags := flags + 1; END_IF;
    IF ok1 THEN flags := flags + 2; END_IF;
    IF ok2 THEN flags := flags + 4; END_IF;
    IF ok3 THEN flags := flags + 8; END_IF;
    IF ok4 THEN flags := flags + 16; END_IF;
    IF ok5 THEN flags := flags + 32; END_IF;
END_PROGRAM

(* ---- o29_muting.st ---- *)
// o29_muting.st — FB_AtcMuting: SafeIn clear n=1..10 & 26..35;
// blocked n=11..25; MutingActive n=11..20 (legit mute) and n=26..30
// (misuse while clear -> MutingBad). flags %QB0: expect 0x1f.
PROGRAM O29
VAR
    flags AT %QB0 : BYTE;
    ok0, ok1, ok2, ok3, ok4 : BOOL;
    mu : FB_AtcMuting;
    n : DINT;
    si, ma : BOOL;
END_VAR
    n := n + 1;
    si := (n <= 10) OR (n >= 26);
    ma := (n >= 11 AND n <= 20) OR (n >= 26 AND n <= 30);
    mu(SafeIn := si, MutingActive := ma, Enable := TRUE,
       CycleTime := 0.1);
    IF n >= 5 AND n <= 10 AND mu.SafeRun AND NOT mu.MuteOut THEN
        ok0 := TRUE;
    END_IF;
    IF n >= 13 AND n <= 19 AND mu.MuteOut AND mu.SafeRun
        AND NOT mu.MutingBad THEN
        ok1 := TRUE;
    END_IF;
    IF n >= 22 AND n <= 25 AND NOT mu.SafeRun AND NOT mu.MuteOut THEN
        ok2 := TRUE;
    END_IF;
    IF n >= 27 AND n <= 30 AND mu.MutingBad AND mu.SafeRun THEN
        ok3 := TRUE;
    END_IF;
    IF n >= 32 AND n <= 35 AND mu.SafeRun AND NOT mu.MuteOut
        AND NOT mu.MutingBad THEN
        ok4 := TRUE;
    END_IF;
    flags := 0;
    IF ok0 THEN flags := flags + 1; END_IF;
    IF ok1 THEN flags := flags + 2; END_IF;
    IF ok2 THEN flags := flags + 4; END_IF;
    IF ok3 THEN flags := flags + 8; END_IF;
    IF ok4 THEN flags := flags + 16; END_IF;
END_PROGRAM

(* ---- o30_valvefb.st ---- *)
// o30_valvefb.st — FB_AtcValveFb: FbDelay=0.5, ct=0.1. Cmd FALSE
// n=11..26 while Fb stays TRUE till n=15 (stuck-open 0.5 s -> Fault
// ~n=15). Cmd=Fb FALSE n=16..26 but Fault latched; Reset n=26.
// Cmd=Fb TRUE again n=28+. flags %QB0: expect 0x3f.
PROGRAM O30
VAR
    flags AT %QB0 : BYTE;
    ok0, ok1, ok2, ok3, ok4, ok5 : BOOL;
    vf : FB_AtcValveFb;
    n : DINT;
    cmd, fb : BOOL;
END_VAR
    n := n + 1;
    cmd := (n <= 10) OR (n >= 27);
    fb := (n <= 15) OR (n >= 28);
    vf(Cmd := cmd, Fb := fb, FbDelay := 0.5, Enable := TRUE,
       CycleTime := 0.1, Reset := (n = 26));
    IF n >= 5 AND n <= 10 AND vf.OK THEN ok0 := TRUE; END_IF;
    IF n >= 12 AND n <= 14 AND NOT vf.OK AND NOT vf.Fault THEN
        ok1 := TRUE;
    END_IF;
    IF n >= 16 AND n <= 20 AND vf.Fault THEN ok2 := TRUE; END_IF;
    IF n >= 21 AND n <= 25 AND NOT vf.OK THEN ok3 := TRUE; END_IF;
    IF n >= 29 AND n <= 33 AND vf.OK AND NOT vf.Fault THEN
        ok4 := TRUE;
    END_IF;
    IF n >= 14 AND n <= 15 AND vf.ET >= 0.3 THEN ok5 := TRUE; END_IF;
    flags := 0;
    IF ok0 THEN flags := flags + 1; END_IF;
    IF ok1 THEN flags := flags + 2; END_IF;
    IF ok2 THEN flags := flags + 4; END_IF;
    IF ok3 THEN flags := flags + 8; END_IF;
    IF ok4 THEN flags := flags + 16; END_IF;
    IF ok5 THEN flags := flags + 32; END_IF;
END_PROGRAM

(* ---- o31_vote.st ---- *)
// o31_vote.st — FB_AtcVote: Band=2.0. Clean triple n=1..10 ->
// median 51. V3=80 n=11..20 -> spread 30 -> Bad, median still 51.
// UseDefault+DefV=45 n=21..25 -> Vout=45 while Bad. Clean again
// n=26..30 -> Bad clears (level, not latched). flags %QB0: 0x1f.
PROGRAM O31
VAR
    flags AT %QB0 : BYTE;
    ok0, ok1, ok2, ok3, ok4 : BOOL;
    vt : FB_AtcVote;
    n : DINT;
    v3 : LREAL;
    ud : BOOL;
END_VAR
    n := n + 1;
    v3 := 52.0;
    IF n >= 11 AND n <= 25 THEN v3 := 80.0; END_IF;
    ud := (n >= 21 AND n <= 25);
    vt(V1 := 50.0, V2 := 51.0, V3 := v3, Band := 2.0,
       UseDefault := ud, DefV := 45.0);
    IF n >= 5 AND n <= 10 AND vt.Vout = 51.0 AND NOT vt.Bad THEN
        ok0 := TRUE;
    END_IF;
    IF n >= 13 AND n <= 19 AND vt.Vout = 51.0 AND vt.Bad
        AND vt.Spread > 25.0 THEN
        ok1 := TRUE;
    END_IF;
    IF n >= 22 AND n <= 25 AND vt.Bad AND vt.Vout = 45.0 THEN
        ok2 := TRUE;
    END_IF;
    IF n >= 27 AND n <= 30 AND vt.Vout = 51.0 AND NOT vt.Bad THEN
        ok3 := TRUE;
    END_IF;
    IF n >= 13 AND n <= 19 AND vt.Spread >= 29.0 AND vt.Spread <= 31.0
    THEN
        ok4 := TRUE;
    END_IF;
    flags := 0;
    IF ok0 THEN flags := flags + 1; END_IF;
    IF ok1 THEN flags := flags + 2; END_IF;
    IF ok2 THEN flags := flags + 4; END_IF;
    IF ok3 THEN flags := flags + 8; END_IF;
    IF ok4 THEN flags := flags + 16; END_IF;
END_PROGRAM

(* ---- o32_loto.st ---- *)
// o32_loto.st — FB_AtcLoto: L2+L5 locked n=11..25 (L2 releases n=21),
// Enable FALSE n=31..35. flags %QB0: expect 0x1f.
PROGRAM O32
VAR
    flags AT %QB0 : BYTE;
    ok0, ok1, ok2, ok3, ok4 : BOOL;
    lo : FB_AtcLoto;
    n : DINT;
    l2, l5 : BOOL;
END_VAR
    n := n + 1;
    l2 := (n >= 11 AND n <= 20);
    l5 := (n >= 11 AND n <= 25);
    lo(L1 := FALSE, L2 := l2, L3 := FALSE, L4 := FALSE,
       L5 := l5, L6 := FALSE, L7 := FALSE, L8 := FALSE,
       Enable := (n < 31 OR n > 35));
    IF n >= 5 AND n <= 10 AND lo.Permit AND lo.LockedCount = 0 THEN
        ok0 := TRUE;
    END_IF;
    IF n >= 13 AND n <= 19 AND NOT lo.Permit AND lo.LockedCount = 2
        AND lo.FirstLock = 2 THEN
        ok1 := TRUE;
    END_IF;
    IF n >= 22 AND n <= 25 AND NOT lo.Permit AND lo.LockedCount = 1
        AND lo.FirstLock = 5 THEN
        ok2 := TRUE;
    END_IF;
    IF n >= 27 AND n <= 30 AND lo.Permit THEN ok3 := TRUE; END_IF;
    IF n >= 32 AND n <= 35 AND NOT lo.Permit THEN ok4 := TRUE; END_IF;
    flags := 0;
    IF ok0 THEN flags := flags + 1; END_IF;
    IF ok1 THEN flags := flags + 2; END_IF;
    IF ok2 THEN flags := flags + 4; END_IF;
    IF ok3 THEN flags := flags + 8; END_IF;
    IF ok4 THEN flags := flags + 16; END_IF;
END_PROGRAM

(* ---- o33_counter.st ---- *)
// o33_counter.st — FB_AtcCounter: Preset=5, ct irrelevant. Up pulses
// n=13,17,21,25,29 (Count->5, AtPreset); Down n=38,44,50 (->2);
// Reset n=55. flags %QB0: expect 0x3f.
PROGRAM O33
VAR
    flags AT %QB0 : BYTE;
    ok0, ok1, ok2, ok3, ok4, ok5 : BOOL;
    ct : FB_AtcCounter;
    n : DINT;
    up, dn : BOOL;
END_VAR
    n := n + 1;
    up := (n >= 11 AND n <= 30) AND (n MOD 4) = 1;
    dn := (n >= 35 AND n <= 52) AND (n MOD 6) = 2;
    ct(Up := up, Down := dn, Preset := 5, Enable := TRUE,
       Reset := (n = 55));
    IF n >= 8 AND n <= 10 AND ct.Count = 0 AND ct.Zero THEN
        ok0 := TRUE;
    END_IF;
    IF n >= 22 AND n <= 24 AND ct.Count = 3 THEN ok1 := TRUE; END_IF;
    IF n >= 30 AND n <= 33 AND ct.AtPreset AND ct.Count = 5 THEN
        ok2 := TRUE;
    END_IF;
    IF n >= 45 AND n <= 49 AND ct.Count = 3 THEN ok3 := TRUE; END_IF;
    IF n >= 51 AND n <= 54 AND ct.Count = 2 AND NOT ct.AtPreset THEN
        ok4 := TRUE;
    END_IF;
    IF n >= 57 AND n <= 60 AND ct.Count = 0 AND ct.Zero THEN
        ok5 := TRUE;
    END_IF;
    flags := 0;
    IF ok0 THEN flags := flags + 1; END_IF;
    IF ok1 THEN flags := flags + 2; END_IF;
    IF ok2 THEN flags := flags + 4; END_IF;
    IF ok3 THEN flags := flags + 8; END_IF;
    IF ok4 THEN flags := flags + 16; END_IF;
    IF ok5 THEN flags := flags + 32; END_IF;
END_PROGRAM

(* ---- o34_ratealarm.st ---- *)
// o34_ratealarm.st — FB_AtcRateAlarm: MaxRate=5, OnDelay=0.5,
// OffDelay=0.3, ct=0.1. PV ramps +2/scan n=11..20 (rate 20 -> Alarm
// ~n=15), holds 70 n=21..30 (clears ~n=23), 72 n=31..35, ramps
// -10/scan n=36..45 (rate -100 -> Alarm ~n=40). flags %QB0: 0x3f.
PROGRAM O34
VAR
    flags AT %QB0 : BYTE;
    ok0, ok1, ok2, ok3, ok4, ok5 : BOOL;
    ra : FB_AtcRateAlarm;
    n : DINT;
    pv : LREAL;
END_VAR
    n := n + 1;
    pv := 50.0;
    IF n >= 11 AND n <= 20 THEN
        pv := 50.0 + 2.0 * DINT_TO_LREAL(n - 10);
    END_IF;
    IF n >= 21 AND n <= 30 THEN pv := 70.0; END_IF;
    IF n >= 31 AND n <= 35 THEN pv := 72.0; END_IF;
    IF n >= 36 AND n <= 45 THEN
        pv := 72.0 - 10.0 * DINT_TO_LREAL(n - 35);
    END_IF;
    IF n >= 46 THEN pv := -28.0; END_IF;
    ra(PV := pv, MaxRate := 5.0, OnDelay := 0.5, OffDelay := 0.3,
       Enable := TRUE, CycleTime := 0.1, Reset := FALSE);
    IF n >= 5 AND n <= 9 AND ra.RateNow = 0.0 AND NOT ra.Alarm THEN
        ok0 := TRUE;
    END_IF;
    IF n >= 12 AND n <= 14 AND ra.RateNow > 15.0 AND NOT ra.Alarm THEN
        ok1 := TRUE;
    END_IF;
    IF n >= 17 AND n <= 20 AND ra.Alarm AND ra.RateNow > 15.0 THEN
        ok2 := TRUE;
    END_IF;
    IF n >= 25 AND n <= 29 AND NOT ra.Alarm THEN ok3 := TRUE; END_IF;
    IF n >= 41 AND n <= 44 AND ra.Alarm AND ra.RateNow < -50.0 THEN
        ok4 := TRUE;
    END_IF;
    IF n = 22 AND ra.Alarm THEN ok5 := TRUE; END_IF;
    flags := 0;
    IF ok0 THEN flags := flags + 1; END_IF;
    IF ok1 THEN flags := flags + 2; END_IF;
    IF ok2 THEN flags := flags + 4; END_IF;
    IF ok3 THEN flags := flags + 8; END_IF;
    IF ok4 THEN flags := flags + 16; END_IF;
    IF ok5 THEN flags := flags + 32; END_IF;
END_PROGRAM

(* ---- o35_delay.st ---- *)
// o35_delay.st — FB_AtcDelay: Delay=0.5 s, ct=0.1 -> 5 samples.
// In=100 pulse at n=3 only; In=50 from n=20. Pulse must appear at
// Out n=8 (5 scans later), step at n=25. Filled once ring >= 5.
// flags %QB0: expect 0x3f.
PROGRAM O35
VAR
    flags AT %QB0 : BYTE;
    ok0, ok1, ok2, ok3, ok4, ok5 : BOOL;
    dl : FB_AtcDelay;
    n : DINT;
    vin : LREAL;
END_VAR
    n := n + 1;
    vin := 0.0;
    IF n = 3 THEN vin := 100.0; END_IF;
    IF n >= 20 THEN vin := 50.0; END_IF;
    dl(In := vin, Delay := 0.5, CycleTime := 0.1, Enable := TRUE,
       Reset := FALSE);
    IF n >= 4 AND n <= 7 AND dl.Out = 0.0 THEN ok0 := TRUE; END_IF;
    IF n = 8 AND dl.Out = 100.0 THEN ok1 := TRUE; END_IF;
    IF n = 9 AND dl.Out = 0.0 THEN ok2 := TRUE; END_IF;
    IF n >= 23 AND n <= 24 AND dl.Out = 0.0 THEN ok3 := TRUE; END_IF;
    IF n >= 26 AND n <= 30 AND dl.Out = 50.0 THEN ok4 := TRUE; END_IF;
    IF n >= 6 AND n <= 10 AND dl.Filled THEN ok5 := TRUE; END_IF;
    flags := 0;
    IF ok0 THEN flags := flags + 1; END_IF;
    IF ok1 THEN flags := flags + 2; END_IF;
    IF ok2 THEN flags := flags + 4; END_IF;
    IF ok3 THEN flags := flags + 8; END_IF;
    IF ok4 THEN flags := flags + 16; END_IF;
    IF ok5 THEN flags := flags + 32; END_IF;
END_PROGRAM

(* ---- o36_ramp.st ---- *)
// o36_ramp.st — FB_AtcRamp: Target=10 always, MaxVel=5, MaxAcc=10,
// ct=0.1. Trapezoid: accel ~5 scans to v=5, cruise, brake ~1.25 u,
// lands Pos=10 Vel=0 Done by ~n=26. flags %QB0: expect 0x3f.
PROGRAM O36
VAR
    flags AT %QB0 : BYTE;
    ok0, ok1, ok2, ok3, ok4, ok5 : BOOL;
    rp : FB_AtcRamp;
    n : DINT;
END_VAR
    n := n + 1;
    rp(Target := 10.0, MaxVel := 5.0, MaxAcc := 10.0,
       Enable := TRUE, CycleTime := 0.1, Reset := FALSE);
    IF n >= 2 AND n <= 4 AND rp.Moving AND rp.Vel > 0.0
        AND rp.Vel < 4.9 THEN
        ok0 := TRUE;
    END_IF;
    IF n >= 10 AND n <= 18 AND rp.Vel = 5.0 AND rp.Moving THEN
        ok1 := TRUE;
    END_IF;
    IF n >= 20 AND n <= 26 AND rp.Vel < 5.0 AND rp.Vel > 0.0
        AND rp.Moving THEN
        ok2 := TRUE;
    END_IF;
    IF n >= 28 AND n <= 40 AND rp.Done AND rp.Pos = 10.0
        AND rp.Vel = 0.0 THEN
        ok3 := TRUE;
    END_IF;
    IF n >= 15 AND n <= 25 AND rp.Pos > 3.0 AND rp.Pos < 10.0 THEN
        ok4 := TRUE;
    END_IF;
    IF n >= 5 AND n <= 9 AND rp.Vel = 5.0 THEN ok5 := TRUE; END_IF;
    flags := 0;
    IF ok0 THEN flags := flags + 1; END_IF;
    IF ok1 THEN flags := flags + 2; END_IF;
    IF ok2 THEN flags := flags + 4; END_IF;
    IF ok3 THEN flags := flags + 8; END_IF;
    IF ok4 THEN flags := flags + 16; END_IF;
    IF ok5 THEN flags := flags + 32; END_IF;
END_PROGRAM

(* ---- o37_ratio.st ---- *)
// o37_ratio.st — FB_AtcRatio: Ratio=0.5, FlowB=10 -> FlowA=6 Total=16;
// Enable off n=11..20 -> FlowA=0 Total=10; FlowB=0 n>=21 -> bias only;
// Bias=2 n>=31 -> FlowA=2. flags %QB0: expect 0x1f.
PROGRAM O37
VAR
    flags AT %QB0 : BYTE;
    ok0, ok1, ok2, ok3, ok4 : BOOL;
    ra : FB_AtcRatio;
    n : DINT;
    fb : LREAL;
    bs : LREAL;
    en : BOOL;
END_VAR
    n := n + 1;
    fb := 10.0;
    IF n >= 21 THEN fb := 0.0; END_IF;
    bs := 1.0;
    IF n >= 31 THEN bs := 2.0; END_IF;
    en := NOT (n >= 11 AND n <= 20);
    ra(FlowB := fb, Ratio := 0.5, Bias := bs, Enable := en);
    IF n >= 5 AND n <= 10 AND ra.FlowA = 6.0 AND ra.Total = 16.0
    THEN
        ok0 := TRUE;
    END_IF;
    IF n >= 13 AND n <= 19 AND ra.FlowA = 0.0 AND ra.Total = 10.0
    THEN
        ok1 := TRUE;
    END_IF;
    IF n >= 23 AND n <= 30 AND ra.FlowA = 1.0 AND ra.Total = 1.0
    THEN
        ok2 := TRUE;
    END_IF;
    IF n >= 32 AND n <= 38 AND ra.FlowA = 2.0 AND ra.Total = 2.0
    THEN
        ok3 := TRUE;
    END_IF;
    IF n = 9 AND ra.FlowA = 6.0 THEN ok4 := TRUE; END_IF;
    flags := 0;
    IF ok0 THEN flags := flags + 1; END_IF;
    IF ok1 THEN flags := flags + 2; END_IF;
    IF ok2 THEN flags := flags + 4; END_IF;
    IF ok3 THEN flags := flags + 8; END_IF;
    IF ok4 THEN flags := flags + 16; END_IF;
END_PROGRAM

(* ---- o38_edge.st ---- *)
// o38_edge.st — FB_AtcEdge: I high n=6..15, pulse n=26, disabled
// pulse n=32 (Enable off n=30..35), I high n=38..42. Edges: rise n=6,
// fall n=16, rise+fall n=26/27, suppressed n=32, rise n=38.
// flags %QB0: expect 0x1f.
PROGRAM O38
VAR
    flags AT %QB0 : BYTE;
    ok0, ok1, ok2, ok3, ok4 : BOOL;
    ed : FB_AtcEdge;
    n : DINT;
    i : BOOL;
    sawQ, sawQN, sawQ2 : BOOL;
END_VAR
    n := n + 1;
    i := (n >= 6 AND n <= 15) OR (n = 26) OR (n = 32)
        OR (n >= 38 AND n <= 42);
    ed(I := i, Enable := NOT (n >= 30 AND n <= 35));
    IF ed.Q THEN sawQ := TRUE; END_IF;
    IF ed.QN THEN sawQN := TRUE; END_IF;
    IF n >= 38 AND ed.Q THEN sawQ2 := TRUE; END_IF;
    IF n >= 8 AND n <= 14 AND NOT ed.Q AND NOT ed.QN THEN
        ok0 := TRUE;
    END_IF;
    IF n >= 20 AND n <= 25 AND NOT ed.Q AND NOT ed.QN THEN
        ok1 := TRUE;
    END_IF;
    IF sawQ THEN ok2 := TRUE; END_IF;
    IF sawQN THEN ok3 := TRUE; END_IF;
    IF sawQ2 THEN ok4 := TRUE; END_IF;
    flags := 0;
    IF ok0 THEN flags := flags + 1; END_IF;
    IF ok1 THEN flags := flags + 2; END_IF;
    IF ok2 THEN flags := flags + 4; END_IF;
    IF ok3 THEN flags := flags + 8; END_IF;
    IF ok4 THEN flags := flags + 16; END_IF;
END_PROGRAM

(* ---- o39_window.st ---- *)
// o39_window.st — FB_AtcWindow: TOD=n. Window 8..20 n<31 (active
// n=8..19); overnight 40..10 n>=31 (active n>=40 or n<10; dead zone
// n=10..39). In=TRUE always. flags %QB0: expect 0x3f.
PROGRAM O39
VAR
    flags AT %QB0 : BYTE;
    ok0, ok1, ok2, ok3, ok4, ok5 : BOOL;
    wn : FB_AtcWindow;
    n : DINT;
    s, e : LREAL;
END_VAR
    n := n + 1;
    s := 8.0; e := 20.0;
    IF n >= 31 THEN s := 40.0; e := 10.0; END_IF;
    wn(In := TRUE, TOD := DINT_TO_LREAL(n), StartT := s, EndT := e);
    IF n >= 3 AND n <= 7 AND NOT wn.Active AND NOT wn.Q THEN
        ok0 := TRUE;
    END_IF;
    IF n >= 10 AND n <= 15 AND wn.Active AND wn.Q THEN ok1 := TRUE;
    END_IF;
    IF n >= 22 AND n <= 28 AND NOT wn.Active THEN ok2 := TRUE; END_IF;
    IF n >= 42 AND n <= 50 AND wn.Active THEN ok3 := TRUE; END_IF;
    IF n >= 60 AND n <= 65 AND wn.Active THEN ok4 := TRUE; END_IF;
    IF n >= 32 AND n <= 38 AND NOT wn.Active THEN ok5 := TRUE; END_IF;
    flags := 0;
    IF ok0 THEN flags := flags + 1; END_IF;
    IF ok1 THEN flags := flags + 2; END_IF;
    IF ok2 THEN flags := flags + 4; END_IF;
    IF ok3 THEN flags := flags + 8; END_IF;
    IF ok4 THEN flags := flags + 16; END_IF;
    IF ok5 THEN flags := flags + 32; END_IF;
END_PROGRAM

(* ---- o40_cam.st ---- *)
// o40_cam.st — FB_AtcCam: trapezoid (0,0)-(10,100)-(20,100)-(30,0),
// X=2n sweep n=1..20. Y interp: X=6->60, plateau 100 for X 10..20,
// X=22->80, X>=30 Sat + Y=0. flags %QB0: expect 0x3f.
PROGRAM O40
VAR
    flags AT %QB0 : BYTE;
    ok0, ok1, ok2, ok3, ok4, ok5 : BOOL;
    cam : FB_AtcCam;
    n : DINT;
    x : LREAL;
END_VAR
    n := n + 1;
    x := DINT_TO_LREAL(n) * 2.0;
    cam.PTS[1].X := 0.0;  cam.PTS[1].Y := 0.0;
    cam.PTS[2].X := 10.0; cam.PTS[2].Y := 100.0;
    cam.PTS[3].X := 20.0; cam.PTS[3].Y := 100.0;
    cam.PTS[4].X := 30.0; cam.PTS[4].Y := 0.0;
    cam(X := x, NPTS := 4, Enable := TRUE);
    IF n = 3 AND cam.Y = 60.0 AND NOT cam.Sat THEN ok0 := TRUE;
    END_IF;
    IF n = 6 AND cam.Y = 100.0 THEN ok1 := TRUE; END_IF;
    IF n = 11 AND cam.Y = 80.0 THEN ok2 := TRUE; END_IF;
    IF n >= 16 AND n <= 20 AND cam.Sat AND cam.Y = 0.0 THEN
        ok3 := TRUE;
    END_IF;
    IF n = 8 AND cam.Y = 100.0 THEN ok4 := TRUE; END_IF;
    IF n >= 17 AND n <= 20 AND cam.Sat THEN ok5 := TRUE; END_IF;
    flags := 0;
    IF ok0 THEN flags := flags + 1; END_IF;
    IF ok1 THEN flags := flags + 2; END_IF;
    IF ok2 THEN flags := flags + 4; END_IF;
    IF ok3 THEN flags := flags + 8; END_IF;
    IF ok4 THEN flags := flags + 16; END_IF;
    IF ok5 THEN flags := flags + 32; END_IF;
END_PROGRAM
